// FB_ModeNodeSpy - test double for the node tree.
//
// A mode node that does nothing except record what the framework did to it:
// how often each Run* method was dispatched, and when in the scan it ran.
// The framework only reaches a node through I_Node and the protected Run*
// methods, so a spy that overrides exactly those sees every call.
FUNCTION_BLOCK FB_ModeNodeSpy EXTENDS FB_ModeNode
VAR_OUTPUT
    nAutomaticCalls : DINT;
    nManualCalls    : DINT;
    nHomingCalls    : DINT;
    nStopCalls      : DINT;
    nScanOrder      : DINT;   // GVL_Test.nScanCounter when this node last ran
END_VAR

// Stamp the scan position, then let FB_ModeNode dispatch by mode as usual.
METHOD PROTECTED OnCyclic
VAR_INPUT
END_VAR
GVL_Test.nScanCounter := GVL_Test.nScanCounter + 1;
nScanOrder := GVL_Test.nScanCounter;
SUPER^.OnCyclic();
END_METHOD

METHOD PROTECTED RunAutomatic
VAR_INPUT
END_VAR
nAutomaticCalls := nAutomaticCalls + 1;
END_METHOD

METHOD PROTECTED RunManual
VAR_INPUT
END_VAR
nManualCalls := nManualCalls + 1;
END_METHOD

METHOD PROTECTED RunHoming
VAR_INPUT
END_VAR
nHomingCalls := nHomingCalls + 1;
END_METHOD

METHOD PROTECTED RunStop
VAR_INPUT
END_VAR
nStopCalls := nStopCalls + 1;
END_METHOD

END_FUNCTION_BLOCK

(* stored: Version 1.1.0.1
   POU FB_ModeNodeSpy: Id {a415b811-aef7-4946-93a9-ade81f586888}, SpecialFunc None
   Method OnCyclic: Id {e0ede19a-c035-435e-afc9-393665eac9fc}
   Method RunAutomatic: Id {4171d4f5-5aa7-4ba2-b744-ad84bc41588a}
   Method RunManual: Id {53e995d9-7e6f-41b4-bb6c-1243224139bf}
   Method RunHoming: Id {c348b9ea-8ba5-4930-bfe7-17cb0edc6d24}
   Method RunStop: Id {b636aa1e-62ce-45fd-b87f-c217d3ac9f67} *)
